(* IEC 61131-3 sources: volt/packages/volt-lsp-iec/test-corpus/bakon-nano/Device/Plc Logic/Application/Library Manager/L_ILMP_LicenseManager, 15 files *)

(* ---- L_ILMP_APPCREDITCONFIGURATION.dut ---- *)
TYPE L_ILMP_APPCREDITCONFIGURATION :
STRUCT
	UDIFASTTOOLBOX : UDINT;
	UDIFASTSERVICES : UDINT;
	UDIFASTUI : UDINT;
	UDIOPCUA : UDINT;
	UDIDEVICEFEATURES : UDINT;
END_STRUCT
END_TYPE

(* ---- L_ILMP_ERROR.dut ---- *)
TYPE L_ILMP_ERROR :
(
	NOERROR := 0,
	NOLICENSEMANAGERAVAILABLE := 16#7100,
	LICENSECONFIGWASALREADYSET := 16#7101,
	WRONGLICENSEMODESELECTED := 16#7102
);
END_TYPE

(* ---- GETBOOLEANPROPERTY.pou ---- *)
FUNCTION GETBOOLEANPROPERTY : BOOL
VAR_INPUT
	STKEY : WSTRING;
END_VAR
END_FUNCTION

(* ---- GETCOMPANY.pou ---- *)
FUNCTION GETCOMPANY : WSTRING
END_FUNCTION

(* ---- GETNUMBERPROPERTY.pou ---- *)
FUNCTION GETNUMBERPROPERTY : DINT
VAR_INPUT
	STKEY : WSTRING;
END_VAR
END_FUNCTION

(* ---- GETTEXTPROPERTY.pou ---- *)
FUNCTION GETTEXTPROPERTY : WSTRING
VAR_INPUT
	STKEY : WSTRING;
END_VAR
END_FUNCTION

(* ---- GETTEXTPROPERTY2.pou ---- *)
FUNCTION GETTEXTPROPERTY2 : POINTER TO WSTRING
VAR_INPUT
	STKEY : WSTRING;
END_VAR
END_FUNCTION

(* ---- GETTITLE.pou ---- *)
FUNCTION GETTITLE : WSTRING
END_FUNCTION

(* ---- GETVERSION.pou ---- *)
FUNCTION GETVERSION : VERSION
END_FUNCTION

(* ---- GETVERSIONPROPERTY.pou ---- *)
FUNCTION GETVERSIONPROPERTY : VERSION
VAR_INPUT
	STKEY : WSTRING;
END_VAR
END_FUNCTION

(* ---- L_ILMP_LICENSECONFIGUPDATEFROMPLC.pou ---- *)
FUNCTION L_ILMP_LICENSECONFIGUPDATEFROMPLC : BOOL
END_FUNCTION

(* ---- L_ILMP_LICENSECONFIGUREMODE.pou ---- *)
FUNCTION L_ILMP_LICENSECONFIGUREMODE : DWORD
VAR_INPUT
	XUPDATE : BOOL;
	DWNEWCONFIGMODE : DWORD;
END_VAR
END_FUNCTION

(* ---- GLOBALTEXTLIST.pou ---- *)
FUNCTION_BLOCK GLOBALTEXTLIST
VAR
	M_TEXTLISTFILE : STRING(255);
	_STNAMESPACE : STRING;
END_VAR
END_FUNCTION_BLOCK

(* ---- L_ILMP_MANAGELICENSECONFIGURATION.pou ---- *)
FUNCTION_BLOCK L_ILMP_MANAGELICENSECONFIGURATION
VAR
	DWCONFIG : DWORD;
	APPLICATIONCREDITINFO : L_IMHP_LM_ApplicationCreditInfo;
	APPCREDITCONFIG : L_IMHP_LM_ApplicationCreditConfiguration;
END_VAR
END_FUNCTION_BLOCK

METHOD INITIALIZE : UDINT
VAR_INPUT
	WMODULETYPE : UINT;
	DWINSTANCE : UDINT;
	PCONNECTOR : POINTER TO IoConfigConnector;
END_VAR
END_METHOD

(* ---- L_ILMP_SETAPPCREDITCONFIGURATION.pou ---- *)
FUNCTION_BLOCK L_ILMP_SETAPPCREDITCONFIGURATION
VAR_INPUT
	XEXECUTE : BOOL;
	SCAPPCREDITCONFIG : L_ILMP_AppCreditConfiguration;
END_VAR
VAR_OUTPUT
	XBUSY : BOOL;
	XDONE : BOOL;
	XERROR : BOOL;
	EERRORID : L_ILMP_Error;
END_VAR
VAR
	XEXECUTEOLD : BOOL;
	DWCONFIG : DWORD;
	XBUSY_INT : BOOL;
	XDONE_INT : BOOL;
	APPLICATIONCREDITINFO : L_IMHP_LM_ApplicationCreditInfo;
	APPCREDITCONFIG : L_IMHP_LM_ApplicationCreditConfiguration;
END_VAR
END_FUNCTION_BLOCK

METHOD ABORT : UDINT
END_METHOD

METHOD EXECUTE : UDINT
END_METHOD
